Staubli VAL3: insertTRAJ.pgx

public program insertTRAJ(string x_sKey, num x_nIndex, string x_sTRAJname, bool& x_bToSave)
  local num l_nIndex
  local num l_i
begin
  if x_nIndex==0 and progTemp:pProgItem[x_sKey].pProgTemplate[x_nIndex].sTRAJname==""
    progTemp:pProgItem[x_sKey].pProgTemplate[x_nIndex].nType=0
    progTemp:pProgItem[x_sKey].pProgTemplate[x_nIndex].sTRAJname=x_sTRAJname
  else
    l_nIndex=x_nIndex+1
    //insert(progTemp:pProgItem[x_sKey].pProgTemplate[x_nIndex+1])
    append(progTemp:pProgItem[x_sKey].pProgTemplate)
    for l_i = size(progTemp:pProgItem[x_sKey].pProgTemplate)-1 to l_nIndex step -1
      call copyPara(x_sKey,l_i-1,l_i)
    endFor
    progTemp:pProgItem[x_sKey].pProgTemplate[x_nIndex+1].nType=0
    progTemp:pProgItem[x_sKey].pProgTemplate[x_nIndex+1].sTRAJname=x_sTRAJname
  endIf

  x_bToSave=true
end
